(* IEC 61131-3 sources: kns-port-domestic/upstream/kns-pump-station/src/POUs/Log/FB_EventLogCsv, 4 files *)

(* ---- FB_EventLogCsv.decl.st ---- *)
// Назначение: выгрузка снимка журнала в CSV через CAA File (SlowTask, PRG_Slow): по фронту xExecute —
//             FILE.Open (MWRITE) → заголовок и строки снимка FB_EventLog по LOG_CSV_LINES_PER_WRITE за один
//             FILE.Write → FILE.Close. Файл — ASCII, «;», CRLF (F_EventCsvLine). Состояние: Writing, затем
//             Done (uiLines строк) или Error (udiError — код FILE.ERROR); держится до следующего фронта.
// Автор:      kr0nsch
// Версия:     0.1.0
// Документ:   docs/DESIGN.md, раздел 9.2; docs/ARCHITECTURE.md, раздел 7
FUNCTION_BLOCK FB_EventLogCsv
VAR_INPUT
    xExecute  : BOOL;               // фронт — начать выгрузку (PRG_Slow: GVL_Log.xExportReq)
    sFileName : STRING(GVL_Const.LOG_PATH_LEN) := GVL_Const.LOG_CSV_FILE;   // относительный путь — каталог рантайма
END_VAR
VAR_IN_OUT
    fbLog : FB_EventLog;            // журнал со снимком (GVL_Log.fbEventLog; TakeSnapshot — MainTask)
END_VAR
VAR_OUTPUT
    eState   : E_LogExportState;    // Idle, Writing, Done, Error
    uiLines  : UINT;                // записано строк данных (без заголовка)
    udiError : UDINT;               // код FILE.ERROR операции с ошибкой; 0 — нет
    xDone    : BOOL;                // файл записан и закрыт
    xError   : BOOL;                // ошибка открытия, записи или закрытия
END_VAR
VAR
    fbOpen    : FILE.Open;
    fbWrite   : FILE.Write;
    fbClose   : FILE.Close;
    xExecPrev : BOOL;               // xExecute прошлого вызова (фронт)
    iStep     : INT;                // шаг выгрузки (STEP_*)
    uiNext    : UINT;               // индекс следующей записи снимка
    xFailed   : BOOL;               // была ошибка записи: после закрытия — Error
    abBuf     : ARRAY[0..GVL_Const.LOG_CSV_BUF_LEN - 1] OF BYTE;   // строки одной операции FILE.Write
    udiBufLen : UDINT;              // байт в abBuf
    stRec     : ST_EventRecord;     // запись снимка
    uiI       : UINT;               // строка порции
END_VAR
VAR CONSTANT
    STEP_IDLE  : INT := 0;
    STEP_OPEN  : INT := 1;
    STEP_WRITE : INT := 2;
    STEP_CLOSE : INT := 3;
    STEP_END   : INT := 4;
    MODE_WRITE : FILE.MODE := FILE.MODE.MWRITE;   // новый файл (существующий перезаписывается)
END_VAR

(* ---- AppendText.method.decl.st ---- *)
// Дописать строку в буфер порции (ASCII-байты без завершающего нуля); не помещается — обрезается по буферу
METHOD PRIVATE AppendText
VAR_INPUT
    sText : STRING(GVL_Const.LOG_CSV_LINE_LEN);
END_VAR
VAR
    pChar : POINTER TO BYTE;       // очередной символ строки
    iI     : INT;                   // номер символа
END_VAR

(* ---- AppendText.method.impl.st ---- *)
pChar := ADR(sText);
FOR iI := 1 TO LEN(sText) DO
    IF udiBufLen < GVL_Const.LOG_CSV_BUF_LEN THEN
        abBuf[udiBufLen] := pChar^;
        udiBufLen := udiBufLen + 1;
    END_IF
    pChar := pChar + 1;
END_FOR

(* ---- FB_EventLogCsv.impl.st ---- *)
// фронт xExecute в покое или после завершения — новая выгрузка
IF xExecute AND NOT xExecPrev AND (iStep = STEP_IDLE OR iStep = STEP_END) THEN
    eState := E_LogExportState.Writing;
    uiLines := 0;
    udiError := 0;
    xDone := FALSE;
    xError := FALSE;
    xFailed := FALSE;
    uiNext := 0;
    iStep := STEP_OPEN;
END_IF
xExecPrev := xExecute;

// шаги: открыть → порции FILE.Write → закрыть
IF iStep = STEP_OPEN THEN
    fbOpen(xExecute := TRUE, sFileName := sFileName, eFileMode := MODE_WRITE, xExclusive := TRUE);
    IF fbOpen.xError THEN
        udiError := TO_UDINT(fbOpen.eError);
        fbOpen(xExecute := FALSE);
        eState := E_LogExportState.Error;
        xError := TRUE;
        iStep := STEP_END;
    ELSIF fbOpen.xDone THEN
        // fbOpen не вызывается до закрытия файла: hFile держится в его выходе
        udiBufLen := 0;
        AppendText(sText := GVL_Const.LOG_CSV_HEADER);
        iStep := STEP_WRITE;
    END_IF
ELSIF iStep = STEP_WRITE THEN
    IF udiBufLen = 0 THEN
        // порция строк снимка
        FOR uiI := 1 TO GVL_Const.LOG_CSV_LINES_PER_WRITE DO
            IF fbLog.GetSnapshotRecord(uiIndex := uiNext, stRecord => stRec) THEN
                AppendText(sText := F_EventCsvLine(stRecord := stRec));
                uiNext := uiNext + 1;
                uiLines := uiLines + 1;
            END_IF
        END_FOR
    END_IF
    IF udiBufLen = 0 THEN
        iStep := STEP_CLOSE;   // снимок выгружен
    ELSE
        fbWrite(xExecute := TRUE, hFile := fbOpen.hFile, pBuffer := ADR(abBuf), szSize := udiBufLen,
                udiTimeOut := GVL_Const.LOG_CSV_TIMEOUT_US);
        IF fbWrite.xError THEN
            udiError := TO_UDINT(fbWrite.eError);
            fbWrite(xExecute := FALSE);
            xFailed := TRUE;
            iStep := STEP_CLOSE;
        ELSIF fbWrite.xDone THEN
            fbWrite(xExecute := FALSE);
            udiBufLen := 0;
        END_IF
    END_IF
ELSIF iStep = STEP_CLOSE THEN
    fbClose(xExecute := TRUE, hFile := fbOpen.hFile);
    IF fbClose.xDone OR fbClose.xError THEN
        IF fbClose.xError AND NOT xFailed THEN
            udiError := TO_UDINT(fbClose.eError);
            xFailed := TRUE;
        END_IF
        fbClose(xExecute := FALSE);
        fbOpen(xExecute := FALSE);
        xError := xFailed;
        xDone := NOT xFailed;
        eState := SEL(xFailed, E_LogExportState.Done, E_LogExportState.Error);
        iStep := STEP_END;
    END_IF
END_IF
